# EPICS substitutions: b-55B2VNC/src/main/epics/PCF0CoreApp/Db/DiamondDetectorDAQ.substitutions
file "DiamondDetectorDAQ.template" {
    pattern { P, PORT }
    { "D1-I2-HWCF:B-0-", "B-0" }
    { "D1-I2-HWCF:B-2-", "B-2" }
}
file "DiamondDetectorDAQ-channel.template" {
    pattern { P, PORT, CH, MIN_LO, MIN_HI }
    { "D1-I2-HWCF:B-0-", "B-0", "0", "-2147483648", "2147483647" }
    { "D1-I2-HWCF:B-0-", "B-0", "1", "-32768", "32767" }
    { "D1-I2-HWCF:B-2-", "B-2", "0", "-2147483648", "2147483647" }
    { "D1-I2-HWCF:B-2-", "B-2", "1", "-32768", "32767" }
}
